ABB RAPID module: FeatureTest.prg

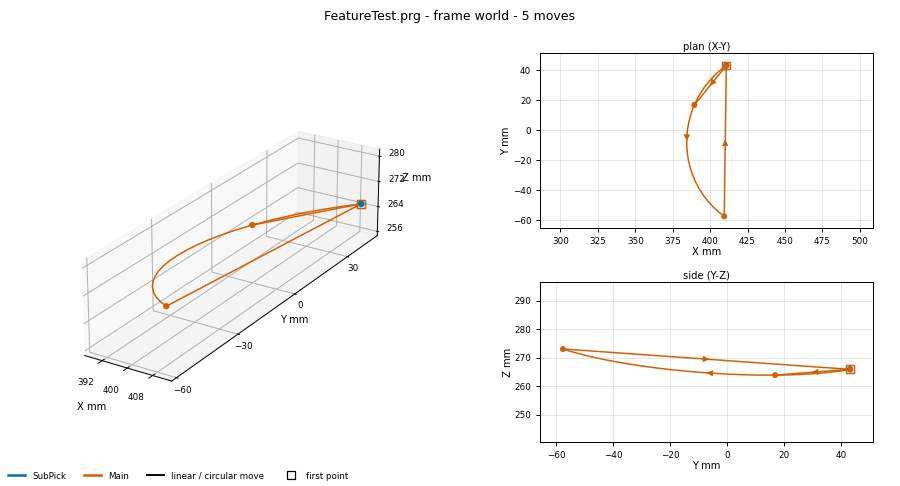
[picture p0: tool path of FeatureTest.prg in frame world, 5 of 7 moves have a stored position in this frame; points joined in program order, loops and branches not executed]
%%%
  VERSION:1
  LANGUAGE:ENGLISH
%%%
MODULE MOD_FeatureTest

    ! -------------------------------
    ! Define customized variables here
    ! ...

	! Tool variables:
	PERS tooldata Tool1 := [TRUE,[[10.000,0.000,120.000],[0.99144486,0.00000000,0.13052619,0.00000001]],[1,[0,0,20],[1,0,0,0],0,0,0.005]];

	! Reference variables:
	PERS wobjdata Frame2 := [FALSE, TRUE, "", [[100.000,-50.000,20.000],[0.96592583,0.00000000,0.00000000,0.25881905]],[[0,0,0],[1,0,0,0]]];

	PROC SubPick()
		ConfJ \On;
		ConfL \Off;
		MoveL [[315.779,-74.668,245.881],[0.09884449,0.01379658,0.99324025,0.05927254],[-1,0,-1,0],[9E+09,9E+09,9E+09,9E+09,9E+09,9E+09]],v300,fine,Tool1 \WObj:=Frame2;
		SetDO D_OUT_7, 1;
	ENDPROC

	PROC Main()
		ConfJ \On;
		ConfL \Off;
		! Program generated by VerticalBot Studio for ABB IRB 120-3/0.6 on 25/10/2026 12:00:00
		! Using nominal kinematics.
		MoveAbsJ [[-10.000000,10.000000,20.000000,30.000000,40.000000,-50.000000],[9E+09,9E+09,9E+09,9E+09,9E+09,9E+09]],v300,z5,Tool1 \WObj:=Frame2;
		MoveL [[315.779,-74.668,245.881],[0.09884449,0.01379658,0.99324025,0.05927254],[-1,0,-1,0],[9E+09,9E+09,9E+09,9E+09,9E+09,9E+09]],v300,z5,Tool1 \WObj:=Frame2;
		MoveC [[284.148,-86.783,243.844],[0.09359571,0.04936652,0.99254150,0.06053239],[-1,0,-1,0],[9E+09,9E+09,9E+09,9E+09,9E+09,9E+09]],[[264.183,-161.234,253.024],[0.11213923,0.13379346,0.98377256,0.04142045],[-1,0,-1,0],[9E+09,9E+09,9E+09,9E+09,9E+09,9E+09]],v300,z5,Tool1 \WObj:=Frame2;
		MoveL [[315.779,-74.668,245.881],[0.09884449,0.01379658,0.99324025,0.05927254],[-1,0,-1,0],[9E+09,9E+09,9E+09,9E+09,9E+09,9E+09]],v50,z0,Tool1 \WObj:=Frame2;
		MoveL [[284.148,-86.783,243.844],[0.09359571,0.04936652,0.99254150,0.06053239],[-1,0,-1,0],[9E+09,9E+09,9E+09,9E+09,9E+09,9E+09]],v300,fine,Tool1 \WObj:=Frame2;
		SetDO D_OUT_3, 1;
		SetDO DO_GRIP, 0;
		WaitDI D_IN_5, 1;
		WaitDI DI_PART, 1, \MaxTime:=2.0;
		WaitTime 0.500;
		! a comment line
		TPWrite "Hello operator";
		MyFunc;
		SetRPM 5000;
		RAW_CODE_LINE
		SubPick;
		Tool1 := [TRUE,[[10.000,0.000,120.000],[0.99144486,0.00000000,0.13052619,0.00000001]],[1,[0,0,20],[1,0,0,0],0,0,0.005]];
		! Attach to Tool 1
		MoveAbsJ [[-10.000000,10.000000,20.000000,30.000000,40.000000,-50.000000],[9E+09,9E+09,9E+09,9E+09,9E+09,9E+09]],v300,fine,Tool1 \WObj:=Frame2;
		STOP;
	ENDPROC

ENDMODULE
